(* IEC 61131-3 sources: vibe-check/src/package-checks/function-metrics/analyzer/fixtures/lizard-1.24.1/st, 3 files *)

(* ---- edge.st ---- *)
FUNCTION reader_sample : INT
VAR_INPUT value : INT; END_VAR
IF value > 0 THEN reader_sample := 1; ELSE reader_sample := 0; END_IF;
END_FUNCTION

(* ---- malformed.st ---- *)
FUNCTION broken : INT
VAR_INPUT value : INT; END_VAR
IF value > 0 THEN

(* ---- normal.st ---- *)
FUNCTION reader_sample : INT
VAR_INPUT value : INT; END_VAR
IF value > 0 THEN reader_sample := 1; ELSE reader_sample := 0; END_IF;
END_FUNCTION
